(*
SPDX-FileCopyrightText: © 2026 Oleksandr Tiutyk <trofimich@gmail.com>
SPDX-License-Identifier: MIT
License: https://opensource.org/license/mit
*)

(*!
<summary>Reports the outcome of a single resetting step in Activity.OnResetting.</summary>
<description>
WORK_IN_PROGRESS keeps the activity in ACTIVE_RESETTING so subsequent Execute calls continue resetting.
WORK_RESET completes resetting, clears stored run diagnostics and transitions the activity to PASSIVE_READY.
</description>
*)

{attribute 'qualified_only'}
{attribute 'strict'}
{attribute 'to_string'}
TYPE ACTIVITY_RESETTING_STATE :
(
	WORK_IN_PROGRESS := 0,
	WORK_RESET
);
END_TYPE

(* stored: Version 1.1.0.1
   DUT ACTIVITY_RESETTING_STATE: Id {45c6b6ea-37c2-4989-9311-5693c5f83e7c} *)
